(*
SPDX-FileCopyrightText: © 2026 Oleksandr Tiutyk <trofimich@gmail.com>
SPDX-License-Identifier: MIT
License: https://opensource.org/license/mit
*)

(*!
<summary>Reports a string length exceeding the limit checked by the caller.</summary>
<description>
The caller detects the error; this type records the supplied diagnostic values without performing the
conversion or validation. Dynamic instances and clones belong to the current task memory manager until
cleanup.
</description>
*)
INTERFACE IStringOverflowException EXTENDS IGeneralException

(*!
<summary>Formats the supplied failure details and propagates this exception.</summary>
<description>
Call in the owning cyclic task, not during FB_init. Captures message, source and timestamps with zero error
code and no inner cause. Input storage is not retained. Allocation failure uses the shared terminal memory
mechanism.
</description>
<param name="actualLength">Actual string length in characters.</param>
<param name="maxLength">Allowed string length in characters.</param>
*)
METHOD Throw
VAR_INPUT
	sourceNamespaceName : STRING;
	sourceClassName : STRING;
	sourcePOUName : STRING;
	sourcePosition : STRING;
	stringName : STRING;
	actualLength : UDINT;
	maxLength : UDINT;
END_VAR
END_METHOD

END_INTERFACE

(* stored: Version 1.1.0.1
   Itf IStringOverflowException: Id {6a53b6ed-b7c4-44c9-9540-6a98d64ca74a}
   Method Throw: Id {370c5aa8-6645-4931-8e8b-bbe194df5099} *)
